(* IEC 61131-3 sources: volt/packages/volt-lsp-iec/test-corpus/CodesysTestProject/Device/Plc Logic/Application/Library Manager/Util, 115 files *)

(* ---- _STATE.dut ---- *)
TYPE _STATE :
(
	UNKNOWN := 0,
	DORMANT,
	STARTING,
	EXECUTING,
	CLEANING,
	DONE,
	ERROR,
	ABORTED,
	RESETTING
);
END_TYPE

(* ---- DATETIME.dut ---- *)
TYPE DATETIME :
STRUCT
	UIYEAR : YEAR;
	UIMONTH : MONTH;
	UIDAY : DAY;
	UIHOUR : HOUR;
	UIMINUTE : MINUTE;
	UISECOND : SECOND;
	UIMILLISECONDS : MILLISECOND;
	EWEEKDAY : WEEKDAY;
END_STRUCT
END_TYPE

(* ---- DAY.dut ---- *)
TYPE DAY : UINT (1..31);
END_TYPE

(* ---- DAYS.dut ---- *)
TYPE DAYS : BYTE;
END_TYPE

(* ---- ERROR.dut ---- *)
TYPE ERROR :
(
	_WRONG_TRANSITION := -1,
	_WRONG_CONFIGURATION := -2,
	NO_ERROR := 0,
	_TIME_OUT := 1,
	WRONG_CONFIGURATION := 2,
	RTC_HIGHRES_NOT_SUPPORTED,
	SYS_TIMEZONE_NOT_SUPPORTED
);
END_TYPE

(* ---- GEN_MODE.dut ---- *)
TYPE GEN_MODE :
(
	TRIANGLE := 0,
	TRIANGLE_POS := 1,
	SAWTOOTH_RISE := 2,
	SAWTOOTH_FALL := 3,
	RECTANGLE := 4,
	SINUS := 5,
	COSINUS := 6,
	SINE := 7,
	COSINE := 8
);
END_TYPE

(* ---- HOUR.dut ---- *)
TYPE HOUR : UINT (0..23);
END_TYPE

(* ---- MILLISECOND.dut ---- *)
TYPE MILLISECOND : UINT (0..999);
END_TYPE

(* ---- MINUTE.dut ---- *)
TYPE MINUTE : UINT (0..59);
END_TYPE

(* ---- MONTH.dut ---- *)
TYPE MONTH : UINT (1..12);
END_TYPE

(* ---- PERIOD.dut ---- *)
TYPE PERIOD :
(
	UNKNOWN := 0,
	STANDARD := 1,
	DAYLIGHT := 2
);
END_TYPE

(* ---- POINT.dut ---- *)
TYPE POINT :
STRUCT
	X : DINT;
	Y : DINT;
END_STRUCT
END_TYPE

(* ---- PT_SIZE.dut ---- *)
TYPE PT_SIZE :
STRUCT
	PSTRING : POINTER TO BYTE;
	UISIZE : UINT;
END_STRUCT
END_TYPE

(* ---- SCHEDULE.dut ---- *)
TYPE SCHEDULE :
STRUCT
	USISWITCH : USINT;
	TODFIRSTON : TIME_OF_DAY;
	TODLASTON : TIME_OF_DAY;
	BYDAYFLAGS : DAYS;
END_STRUCT
END_TYPE

(* ---- SECOND.dut ---- *)
TYPE SECOND : MINUTE;
END_TYPE

(* ---- SEGMENT.dut ---- *)
TYPE SEGMENT :
STRUCT
	SNAME : TZ_NAME;
	DTDATE : DateTime;
	IBIAS : INT;
END_STRUCT
END_TYPE

(* ---- TIMEZONE.dut ---- *)
TYPE TIMEZONE :
STRUCT
	IBIAS : INT;
	ASGPERIOD : ARRAY [1..2] OF Segment;
END_STRUCT
END_TYPE

(* ---- TZ_NAME.dut ---- *)
TYPE TZ_NAME : STRING(32);
END_TYPE

(* ---- WEEK.dut ---- *)
TYPE WEEK : UINT (1..53);
END_TYPE

(* ---- WEEKDAY.dut ---- *)
TYPE WEEKDAY :
(
	UNKNOWN := 0,
	MONDAY := 1,
	TUESDAY := 2,
	WEDNESDAY := 3,
	THURSDAY := 4,
	FRIDAY := 5,
	SATURDAY := 6,
	SUNDAY := 7
);
END_TYPE

(* ---- YEAR.dut ---- *)
TYPE YEAR : UINT (0..2106);
END_TYPE

(* ---- CONSTANTS.gvl ---- *)
VAR_GLOBAL
	GC_ULISECONDSINDAY : ULINT := (ANY_TO_ULINT(TIME#1440m0s0ms) / 1000);
	GC_AUSIWEEKDAY : ARRAY [0..11] OF USINT := [0, 3, 3, 6, 1, 4, 6, 2, 5, 0, 3, 5];
	GC_AUSIDAYSINMONTH : ARRAY [0..11] OF USINT := [31, 28, 31, 30, 31, 30, 31, 31, 30, 31, 30, 31];
	GC_AUIDAYSINYEAR : ARRAY [0..11] OF UINT := [0, 31, 59, 90, 120, 151, 181, 212, 243, 273, 304, 334];
	GC_DWSWITCHMASK : ARRAY [0..31] OF DWORD := [16#1, 16#2, 16#4, 16#8, 16#10, 16#20, 16#40, 16#80, 16#100, 16#200, 16#400, 16#800, 16#1000, 16#2000, 16#4000, 16#8000, 16#10000, 16#20000, 16#40000, 16#80000, 16#100000, 16#200000, 16#400000, 16#800000, 16#1000000, 16#2000000, 16#4000000, 16#8000000, 16#10000000, 16#20000000, 16#40000000, 16#80000000];
	GC_BYDAYMASK : ARRAY [0..7] OF DAYS := [DAY_FLAGS.EVERY_DAY, DAY_FLAGS.MONDAY, DAY_FLAGS.TUESDAY, DAY_FLAGS.WEDNESDAY, DAY_FLAGS.THURSDAY, DAY_FLAGS.FRIDAY, DAY_FLAGS.SATURDAY, DAY_FLAGS.SUNDAY];
END_VAR

(* ---- DAY_FLAGS.gvl ---- *)
VAR_GLOBAL
	EVERY_DAY : DAYS := 0;
	WORKING_DAYS : DAYS := 31;
	WEEKEND : DAYS := 96;
	MONDAY : DAYS := 1;
	TUESDAY : DAYS := 2;
	WEDNESDAY : DAYS := 4;
	THURSDAY : DAYS := 8;
	FRIDAY : DAYS := 16;
	SATURDAY : DAYS := 32;
	SUNDAY : DAYS := 64;
END_VAR

(* ---- GLOBALS.gvl ---- *)
VAR_GLOBAL
	G_DTPDATETIMEPROVIDER : DateTimeProvider;
END_VAR

(* ---- GVL_CONST.gvl ---- *)
VAR_GLOBAL
	UIBLOCKSIZEENCODED : UINT := REAL_TO_UINT((TextBlockSize.iBlockSize + (TextBlockSize.iBlockSize * 0.35)));
END_VAR

(* ---- TEXTBLOCKSIZE.gvl ---- *)
VAR_GLOBAL
	IBLOCKSIZE : INT := 22800;
END_VAR

(* ---- TSW.gvl ---- *)
VAR_GLOBAL
	GC_TZTIMEZONECET : TimeZone := STRUCT(iBias := 60, asgPeriod := [STRUCT(sName := 'CET', dtDate := STRUCT(uiMonth := 10, eWeekday := WEEKDAY.SUNDAY, uiDay := 5, uiHour := 3)), STRUCT(sName := 'CEST', dtDate := STRUCT(uiMonth := 3, eWeekday := WEEKDAY.SUNDAY, uiDay := 5, uiHour := 2), iBias := 60)]);
	GC_TZTIMEZONEUTC : TimeZone := STRUCT(asgPeriod := [STRUCT(sName := 'UTC')]);
END_VAR

(* ---- _IACTIONCONTROLLER.itf ---- *)
INTERFACE _IACTIONCONTROLLER
END_INTERFACE

METHOD CONTROLCLEANUPACTION
VAR_INPUT
	ITFCLEANUPACTIONPROVIDER : _ICleanupActionProvider;
	XABORTPROPOSED : BOOL;
	IERRORIDPROPOSED : INT;
END_VAR
VAR_OUTPUT
	XCOMPLETE : BOOL;
	XABORT : BOOL;
	IERRORID : INT;
END_VAR
END_METHOD

METHOD CONTROLCYCLICACTION
VAR_INPUT
	ITFCYCLICACTIONPROVIDER : _ICyclicActionProvider;
	ITFTIMINGCONTROLLER : _ITimingController;
END_VAR
VAR_OUTPUT
	XCOMPLETE : BOOL;
	IERRORID : INT;
END_VAR
END_METHOD

METHOD CONTROLEXITACTION
VAR_INPUT
	ITFEXITACTIONPROVIDER : _IExitActionProvider;
	XAFTERCLEANUP : BOOL;
	XINCOPYCODE : BOOL;
END_VAR
END_METHOD

METHOD CONTROLRESETACTION
VAR_INPUT
	ITFRESETACTIONPROVIDER : _IResetActionProvider;
END_VAR
VAR_OUTPUT
	XCOMPLETE : BOOL;
END_VAR
END_METHOD

METHOD CONTROLSTARTACTION
VAR_INPUT
	ITFSTARTACTIONPROVIDER : _IStartActionProvider;
END_VAR
VAR_OUTPUT
	XCOMPLETE : BOOL;
	IERRORID : INT;
END_VAR
END_METHOD

(* ---- _IACTIONPROVIDER.itf ---- *)
INTERFACE _IACTIONPROVIDER
END_INTERFACE

(* ---- _IBEHAVIOURMODEL.itf ---- *)
INTERFACE _IBEHAVIOURMODEL
END_INTERFACE

METHOD ABORTMODEL : ERROR
VAR_INPUT
	XCOMMIT : BOOL;
END_VAR
END_METHOD

METHOD GETMODELSTATE
VAR_INPUT
	XCOMMIT : BOOL;
END_VAR
VAR_OUTPUT
	XDONE : BOOL;
	XBUSY : BOOL;
	XERROR : BOOL;
	XABORTED : BOOL;
	IERRORID : INT;
	ESTATE : _STATE;
END_VAR
END_METHOD

METHOD RESETMODEL : ERROR
VAR_INPUT
	XCOMMIT : BOOL;
END_VAR
END_METHOD

METHOD STARTMODEL : ERROR
VAR_INPUT
	XCOMMIT : BOOL;
END_VAR
END_METHOD

(* ---- _ICLEANUPACTIONPROVIDER.itf ---- *)
INTERFACE _ICLEANUPACTIONPROVIDER
END_INTERFACE

METHOD CLEANUPACTION
VAR_INPUT
	XABORTPROPOSED : BOOL;
	IERRORIDPROPOSED : INT;
END_VAR
VAR_OUTPUT
	XCOMPLETE : BOOL;
	XABORT : BOOL;
	IERRORID : INT;
END_VAR
END_METHOD

(* ---- _ICONFIGURATIONPROVIDER.itf ---- *)
INTERFACE _ICONFIGURATIONPROVIDER
END_INTERFACE

METHOD GETCONFIGURATION
VAR_OUTPUT
	XLEVELCONTROLLED : BOOL;
	XTIMINGCONTROLLED : BOOL;
	XTIMELIMITED : BOOL;
	XTIMEOUTCONSTRAINT : BOOL;
	XABORTABLE : BOOL;
	XEDGETRIGGERED : BOOL;
	XHASCONTINUOUSBEHAVIOUR : BOOL;
	XSUPPORTSEXITACTION : BOOL;
END_VAR
END_METHOD

(* ---- _ICONFIGURATIONPROVIDER2.itf ---- *)
INTERFACE _ICONFIGURATIONPROVIDER2
END_INTERFACE

METHOD GETCONFIGURATION2
VAR_OUTPUT
	XLEVELCONTROLLED : BOOL;
	XTIMINGCONTROLLED : BOOL;
	XTIMELIMITED : BOOL;
	XTIMEOUTCONSTRAINT : BOOL;
	XABORTABLE : BOOL;
	XEDGETRIGGERED : BOOL;
	XHASCONTINUOUSBEHAVIOUR : BOOL;
	XSUPPORTSEXITACTION : BOOL;
	XSUPPORTSSAMPLEACTION : BOOL;
END_VAR
END_METHOD

(* ---- _ICYCLICACTIONPROVIDER.itf ---- *)
INTERFACE _ICYCLICACTIONPROVIDER
END_INTERFACE

METHOD CYCLICACTION
VAR_INPUT
	ITFTIMINGCONTROLLER : _ITimingController;
END_VAR
VAR_OUTPUT
	XCOMPLETE : BOOL;
	IERRORID : INT;
END_VAR
END_METHOD

(* ---- _IEXITACTIONPROVIDER.itf ---- *)
INTERFACE _IEXITACTIONPROVIDER
END_INTERFACE

METHOD EXITACTION
VAR_INPUT
	XAFTERCLEANUP : BOOL;
	XINCOPYCODE : BOOL;
END_VAR
END_METHOD

(* ---- _IHASCONTINUOUSBEHAVIOUR.itf ---- *)
INTERFACE _IHASCONTINUOUSBEHAVIOUR
END_INTERFACE

(* ---- _ILEVELCONTROLLED.itf ---- *)
INTERFACE _ILEVELCONTROLLED
END_INTERFACE

(* ---- _IRESETACTIONPROVIDER.itf ---- *)
INTERFACE _IRESETACTIONPROVIDER
END_INTERFACE

METHOD RESETACTION
VAR_OUTPUT
	XCOMPLETE : BOOL;
END_VAR
END_METHOD

(* ---- _ISTARTACTIONPROVIDER.itf ---- *)
INTERFACE _ISTARTACTIONPROVIDER
END_INTERFACE

METHOD STARTACTION
VAR_OUTPUT
	XCOMPLETE : BOOL;
	IERRORID : INT;
END_VAR
END_METHOD

(* ---- _ITIMINGCONTROLLER.itf ---- *)
INTERFACE _ITIMINGCONTROLLER
END_INTERFACE

METHOD CONTROLLERCHECKTIMING
VAR_OUTPUT
	XTIMEOUT : BOOL;
	XTIMELIMIT : BOOL;
END_VAR
END_METHOD

METHOD STARTINVOCATIONTIMER
END_METHOD

METHOD STARTOPERATIONTIMER
END_METHOD

(* ---- IDATETIMEPROVIDER.itf ---- *)
INTERFACE IDATETIMEPROVIDER
END_INTERFACE

METHOD GETDATETIME : ULINT
VAR_OUTPUT
	EERRORID : ERROR;
END_VAR
END_METHOD

(* ---- ITIMESWITCH.itf ---- *)
INTERFACE ITIMESWITCH
END_INTERFACE

(* ---- BASE64.pou ---- *)
FUNCTION BASE64 : PT_SIZE
VAR_INPUT
	TEXTTOENCODE : PT_SIZE;
	ISLASTBLOCK : BOOL;
	PBYERROR : POINTER TO BYTE;
END_VAR
END_FUNCTION

(* ---- BCD_TO_BYTE.pou ---- *)
FUNCTION BCD_TO_BYTE : BYTE
VAR_INPUT
	B : BYTE;
END_VAR
END_FUNCTION

(* ---- BCD_TO_DWORD.pou ---- *)
FUNCTION BCD_TO_DWORD : DWORD
VAR_INPUT
	X : DWORD;
END_VAR
END_FUNCTION

(* ---- BCD_TO_INT.pou ---- *)
FUNCTION BCD_TO_INT : INT
VAR_INPUT
	B : BYTE;
END_VAR
END_FUNCTION

(* ---- BCD_TO_WORD.pou ---- *)
FUNCTION BCD_TO_WORD : WORD
VAR_INPUT
	W : WORD;
END_VAR
END_FUNCTION

(* ---- BYTE_TO_BCD.pou ---- *)
FUNCTION BYTE_TO_BCD : BYTE
VAR_INPUT
	B : BYTE;
END_VAR
END_FUNCTION

(* ---- BYTE_TO_GRAY.pou ---- *)
FUNCTION BYTE_TO_GRAY : BYTE
VAR_INPUT
	B : BYTE;
END_VAR
END_FUNCTION

(* ---- BYTE_TO_HEXINASCII.pou ---- *)
FUNCTION BYTE_TO_HEXINASCII : WORD
VAR_INPUT
	B : BYTE;
END_VAR
END_FUNCTION

(* ---- COMBINEDATETIME.pou ---- *)
FUNCTION COMBINEDATETIME : ULINT
VAR_INPUT
	DATDATE : DATE;
	TODTIME : TIME_OF_DAY;
END_VAR
VAR_OUTPUT
	EERRORID : ERROR := ERROR.NO_ERROR;
END_VAR
END_FUNCTION

(* ---- CONVERTDATETIME.pou ---- *)
FUNCTION CONVERTDATETIME : ULINT
VAR_INPUT
	UIYEAR : YEAR;
END_VAR
VAR_OUTPUT
	EERRORID : ERROR;
END_VAR
VAR_IN_OUT
	DTDATETIME : DateTime;
END_VAR
END_FUNCTION

(* ---- DATETIMEFROMWEEK.pou ---- *)
FUNCTION DATETIMEFROMWEEK : ULINT
VAR_INPUT
	UIYEAR : YEAR;
	UIWEEK : WEEK;
	EWEEKDAY : WEEKDAY;
END_VAR
VAR_OUTPUT
	EERRORID : ERROR;
END_VAR
END_FUNCTION

(* ---- DAYOFWEEK.pou ---- *)
FUNCTION DAYOFWEEK : WEEKDAY
VAR_INPUT
	DATDATE : DATE;
END_VAR
VAR_OUTPUT
	EERRORID : ERROR := ERROR.NO_ERROR;
END_VAR
END_FUNCTION

(* ---- DWORD_TO_BCD.pou ---- *)
FUNCTION DWORD_TO_BCD : DWORD
VAR_INPUT
	X : DWORD;
END_VAR
END_FUNCTION

(* ---- DWORD_TO_GRAY.pou ---- *)
FUNCTION DWORD_TO_GRAY : DWORD
VAR_INPUT
	X : DWORD;
END_VAR
END_FUNCTION

(* ---- EXTRACT.pou ---- *)
FUNCTION EXTRACT : BOOL
VAR_INPUT
	X : DWORD;
	N : BYTE;
END_VAR
END_FUNCTION

(* ---- EXTRACTYEARMONTHDAY.pou ---- *)
FUNCTION EXTRACTYEARMONTHDAY : ERROR
VAR_INPUT
	ULIDATETIME : ULINT;
END_VAR
VAR_OUTPUT
	UIYEAR : YEAR;
	UIMONTH : MONTH;
	UIDAY : DAY;
END_VAR
END_FUNCTION

(* ---- GETBIT.pou ---- *)
FUNCTION GETBIT : BOOL
VAR_INPUT
	X : LWORD;
	N : BYTE;
END_VAR
END_FUNCTION

(* ---- GETDATETIME.pou ---- *)
FUNCTION GETDATETIME : ULINT
VAR_OUTPUT
	EERRORID : ERROR;
END_VAR
END_FUNCTION

(* ---- GETLIBVERSION.pou ---- *)
FUNCTION GETLIBVERSION : VERSION
END_FUNCTION

(* ---- GETLIBVERSIONNUMBER.pou ---- *)
FUNCTION GETLIBVERSIONNUMBER : DWORD
END_FUNCTION

(* ---- GETLOCALDATETIME.pou ---- *)
FUNCTION GETLOCALDATETIME : ULINT
VAR_OUTPUT
	EERRORID : ERROR;
END_VAR
VAR_IN_OUT
	TZTIMEZONE : TimeZone;
END_VAR
END_FUNCTION

(* ---- GETTIMESTAMPSDIFFERENCE.pou ---- *)
FUNCTION GETTIMESTAMPSDIFFERENCE : ERROR
VAR_INPUT
	ULIDATETIMEFIRST : ULINT;
	ULIDATETIMESECOND : ULINT;
END_VAR
VAR_OUTPUT
	ULIDAYS : ULINT;
	UIHOURS : HOUR;
	UIMINUTES : MINUTE;
	UISECONDS : SECOND;
	UIMILLISECONDS : MILLISECOND;
END_VAR
END_FUNCTION

(* ---- GRAY_TO_BYTE.pou ---- *)
FUNCTION GRAY_TO_BYTE : BYTE
VAR_INPUT
	B : BYTE;
END_VAR
END_FUNCTION

(* ---- GRAY_TO_DWORD.pou ---- *)
FUNCTION GRAY_TO_DWORD : DWORD
VAR_INPUT
	X : DWORD;
END_VAR
END_FUNCTION

(* ---- GRAY_TO_WORD.pou ---- *)
FUNCTION GRAY_TO_WORD : WORD
VAR_INPUT
	W : WORD;
END_VAR
END_FUNCTION

(* ---- HEXINASCII_TO_BYTE.pou ---- *)
FUNCTION HEXINASCII_TO_BYTE : BYTE
VAR_INPUT
	W : WORD;
END_VAR
END_FUNCTION

(* ---- INT_TO_BCD.pou ---- *)
FUNCTION INT_TO_BCD : BYTE
VAR_INPUT
	I : INT;
END_VAR
END_FUNCTION

(* ---- ISLEAPYEAR.pou ---- *)
FUNCTION ISLEAPYEAR : BOOL
VAR_INPUT
	UIYEAR : YEAR;
END_VAR
VAR_OUTPUT
	EERRORID : ERROR := ERROR.NO_ERROR;
END_VAR
END_FUNCTION

(* ---- ISLIBRELEASED.pou ---- *)
FUNCTION ISLIBRELEASED : BOOL
END_FUNCTION

(* ---- JOINDATETIME.pou ---- *)
FUNCTION JOINDATETIME : ULINT
VAR_INPUT
	UIYEAR : YEAR;
	UIMONTH : MONTH;
	UIDAY : DAY;
	UIHOUR : HOUR;
	UIMINUTE : MINUTE;
	UISECOND : SECOND;
	UIMILLISECONDS : MILLISECOND;
END_VAR
VAR_OUTPUT
	EERRORID : ERROR := ERROR.NO_ERROR;
END_VAR
END_FUNCTION

(* ---- JOINYEARMONTHDAY.pou ---- *)
FUNCTION JOINYEARMONTHDAY : ULINT
VAR_INPUT
	UIYEAR : YEAR;
	UIMONTH : MONTH;
	UIDAY : DAY;
END_VAR
VAR_OUTPUT
	EERRORID : ERROR := ERROR.NO_ERROR;
END_VAR
END_FUNCTION

(* ---- LASTWEEKOFYEAR.pou ---- *)
FUNCTION LASTWEEKOFYEAR : Week
VAR_INPUT
	UIYEAR : YEAR;
END_VAR
VAR_OUTPUT
	EERRORID : ERROR;
END_VAR
END_FUNCTION

(* ---- LEAPYEARS.pou ---- *)
FUNCTION LEAPYEARS : UINT
VAR_INPUT
	UISTARTYEAR : YEAR;
	UIENDYEAR : YEAR;
END_VAR
VAR_OUTPUT
	EERRORID : ERROR;
END_VAR
END_FUNCTION

(* ---- LOCALDATETIME.pou ---- *)
FUNCTION LOCALDATETIME : ULINT
VAR_INPUT
	ULIDATETIME : ULINT;
END_VAR
VAR_OUTPUT
	EERRORID : ERROR;
	EPERIOD : PERIOD;
END_VAR
VAR_IN_OUT
	TZTIMEZONE : TimeZone;
END_VAR
END_FUNCTION

(* ---- PACK.pou ---- *)
FUNCTION PACK : BYTE
VAR_INPUT
	B0 : BOOL;
	B1 : BOOL;
	B2 : BOOL;
	B3 : BOOL;
	B4 : BOOL;
	B5 : BOOL;
	B6 : BOOL;
	B7 : BOOL;
END_VAR
END_FUNCTION

(* ---- PUTBIT.pou ---- *)
FUNCTION PUTBIT : DWORD
VAR_INPUT
	X : DWORD;
	N : BYTE;
	B : BOOL;
END_VAR
END_FUNCTION

(* ---- SEPARATEDATETIME.pou ---- *)
FUNCTION SEPARATEDATETIME : ERROR
VAR_INPUT
	ULIDATETIME : ULINT;
END_VAR
VAR_OUTPUT
	EWEEKDAY : WEEKDAY;
	DATDATE : DATE;
	TODTIME : TIME_OF_DAY;
END_VAR
END_FUNCTION

(* ---- SETBIT.pou ---- *)
FUNCTION SETBIT : BOOL
VAR_INPUT
	X : __SYSTEM.AnyType;
	N : BYTE;
	B : BOOL;
END_VAR
END_FUNCTION

(* ---- SPLITDATETIME.pou ---- *)
FUNCTION SPLITDATETIME : ERROR
VAR_INPUT
	ULIDATETIME : ULINT;
END_VAR
VAR_OUTPUT
	UIYEAR : YEAR;
	UIMONTH : MONTH;
	UIDAY : DAY;
	UIHOUR : HOUR;
	UIMINUTE : MINUTE;
	UISECOND : SECOND;
	UIMILLISECONDS : MILLISECOND;
	EWEEKDAY : WEEKDAY;
END_VAR
END_FUNCTION

(* ---- SWITCHBIT.pou ---- *)
FUNCTION SWITCHBIT : DWORD
VAR_INPUT
	X : DWORD;
	N : BYTE;
END_VAR
END_FUNCTION

(* ---- WEEKOFYEAR.pou ---- *)
FUNCTION WEEKOFYEAR : ERROR
VAR_INPUT
	ULIDATETIME : ULINT;
END_VAR
VAR_OUTPUT
	UIYEAR : YEAR;
	UIWEEK : WEEK;
	EWEEKDAY : WEEKDAY;
END_VAR
END_FUNCTION

(* ---- WORD_AS_STRING.pou ---- *)
FUNCTION WORD_AS_STRING : STRING(2)
VAR_INPUT
	W : WORD;
	ORDER : BOOL;
END_VAR
END_FUNCTION

(* ---- WORD_TO_BCD.pou ---- *)
FUNCTION WORD_TO_BCD : WORD
VAR_INPUT
	W : WORD;
END_VAR
END_FUNCTION

(* ---- WORD_TO_GRAY.pou ---- *)
FUNCTION WORD_TO_GRAY : WORD
VAR_INPUT
	W : WORD;
END_VAR
END_FUNCTION

(* ---- _BEHAVIOURMODEL.pou ---- *)
FUNCTION_BLOCK _BEHAVIOURMODEL
VAR_INPUT
	ITFACTIONPROVIDER : _IActionProvider;
	ITFTIMINGCONTROLLER : _ITimingController;
	XCONTROL : BOOL;
	XABORT : BOOL;
	UDITIMELIMIT : UDINT;
	UDITIMEOUT : UDINT;
END_VAR
VAR_OUTPUT
	XDONE : BOOL;
	XBUSY : BOOL;
	XERROR : BOOL;
	XABORTED : BOOL;
	IERRORID : INT;
	ESTATE : _STATE;
	EINTERNALERRORID : ERROR;
END_VAR
VAR
	_ITFACTIONPROVIDER : _IActionProvider;
	_ITFACTIONCONTROLLER : _IActionController;
	_XLEVELCONTROLLED : BOOL;
	_XTIMINGCONTROLLED : BOOL;
	_XTIMELIMITED : BOOL;
	_XTIMEOUTCONSTRAINT : BOOL;
	_XABORTABLE : BOOL;
	_XEDGETRIGGERED : BOOL;
	_XHASCONTINUOUSBEHAVIOUR : BOOL;
	_XSUPPORTSEXITACTION : BOOL;
	_XSUPPORTSSAMPLEACTION : BOOL;
	_XRESETREQUEST : BOOL;
	_XABORTPROPOSED : BOOL;
	_IERRORIDPROPOSED : INT;
	_XFIRSTHANDLESTARTINGSTATECALL : BOOL;
	_XLASTAGAIN : BOOL;
	_ITFSTARTACTIONPROVIDER : _IStartActionProvider;
	_ITFCYCLICACTIONPROVIDER : _ICyclicActionProvider;
	_ITFCLEANUPACTIONPROVIDER : _ICleanupActionProvider;
	_ITFEXITACTIONPROVIDER : _IExitActionProvider;
	_ITFRESETACTIONPROVIDER : _IResetActionProvider;
	ACTIONCONTROLLER : _IActionController;
	MODELTIMELIMIT : UDINT;
	MODELTIMEOUT : UDINT;
END_VAR
END_FUNCTION_BLOCK

METHOD _CHECKABORTCONDITION : BOOL
END_METHOD

METHOD _CHECKPARAMETER
VAR_OUTPUT
	EERRORID : ERROR;
END_VAR
END_METHOD

METHOD _CHECKTIMEOUTCONDITION
END_METHOD

METHOD _EXECUTE
VAR_OUTPUT
	EERRORID : ERROR := ERROR.NO_ERROR;
END_VAR
END_METHOD

METHOD _RESETACTION
END_METHOD

METHOD ABORTMODEL : ERROR
VAR_INPUT
	XCOMMIT : BOOL;
END_VAR
END_METHOD

METHOD GETCONFIGURATION
VAR_OUTPUT
	XLEVELCONTROLLED : BOOL;
	XTIMINGCONTROLLED : BOOL;
	XTIMELIMITED : BOOL;
	XTIMEOUTCONSTRAINT : BOOL;
	XABORTABLE : BOOL;
	XEDGETRIGGERED : BOOL;
	XHASCONTINUOUSBEHAVIOUR : BOOL;
	XSUPPORTSEXITACTION : BOOL;
END_VAR
END_METHOD

METHOD GETCONFIGURATION2
VAR_OUTPUT
	XLEVELCONTROLLED : BOOL;
	XTIMINGCONTROLLED : BOOL;
	XTIMELIMITED : BOOL;
	XTIMEOUTCONSTRAINT : BOOL;
	XABORTABLE : BOOL;
	XEDGETRIGGERED : BOOL;
	XHASCONTINUOUSBEHAVIOUR : BOOL;
	XSUPPORTSEXITACTION : BOOL;
	XSUPPORTSSAMPLEACTION : BOOL;
END_VAR
END_METHOD

METHOD GETMODELSTATE
VAR_INPUT
	XCOMMIT : BOOL;
END_VAR
VAR_OUTPUT
	XDONE : BOOL;
	XBUSY : BOOL;
	XERROR : BOOL;
	XABORTED : BOOL;
	IERRORID : INT;
	ESTATE : _STATE;
END_VAR
END_METHOD

METHOD RESETMODEL : ERROR
VAR_INPUT
	XCOMMIT : BOOL;
END_VAR
END_METHOD

METHOD STARTMODEL : ERROR
VAR_INPUT
	XCOMMIT : BOOL;
END_VAR
END_METHOD

METHOD _HANDLEABORTEDSTATE
VAR_OUTPUT
	XAGAIN : BOOL;
END_VAR
END_METHOD

METHOD _HANDLECLEANINGSTATE
VAR_OUTPUT
	XAGAIN : BOOL;
END_VAR
END_METHOD

METHOD _HANDLEDONESTATE
VAR_OUTPUT
	XAGAIN : BOOL;
END_VAR
END_METHOD

METHOD _HANDLEDORMANTSTATE
VAR_OUTPUT
	XAGAIN : BOOL;
END_VAR
END_METHOD

METHOD _HANDLEERRORSTATE
VAR_OUTPUT
	XAGAIN : BOOL;
END_VAR
END_METHOD

METHOD _HANDLEEXECUTINGSTATE
VAR_OUTPUT
	XAGAIN : BOOL;
END_VAR
END_METHOD

METHOD _HANDLERESETTINGSTATE
VAR_OUTPUT
	XAGAIN : BOOL;
END_VAR
END_METHOD

METHOD _HANDLESTARTINGSTATE
VAR_OUTPUT
	XAGAIN : BOOL;
	IERRORID : INT;
END_VAR
END_METHOD

METHOD _STATEMACHINE : ERROR
END_METHOD

(* ---- _LCONC.pou ---- *)
FUNCTION_BLOCK _LCONC
VAR_INPUT
	XENABLE : BOOL;
END_VAR
VAR_OUTPUT
	XBUSY : BOOL;
	XERROR : BOOL;
END_VAR
VAR
	_MODEL : _BehaviourModel := STRUCT(itfActionProvider := THIS^, itfTimingController := 0);
	ACTIONCONTROLLER : _IActionController;
	MODELTIMELIMIT : UDINT;
	MODELTIMEOUT : UDINT;
END_VAR
END_FUNCTION_BLOCK

METHOD FB_EXIT : BOOL
VAR_INPUT
	BINCOPYCODE : BOOL;
END_VAR
END_METHOD

METHOD _EXECUTE
VAR_OUTPUT
	EERRORID : ERROR;
END_VAR
END_METHOD

METHOD CLEANUPACTION
VAR_INPUT
	XABORTPROPOSED : BOOL;
	IERRORIDPROPOSED : INT;
END_VAR
VAR_OUTPUT
	XCOMPLETE : BOOL := TRUE;
	XABORT : BOOL := xAbortProposed;
	IERRORID : INT := iErrorIDProposed;
END_VAR
END_METHOD

METHOD CYCLICACTION
VAR_INPUT
	ITFTIMINGCONTROLLER : _ITimingController;
END_VAR
VAR_OUTPUT
	XCOMPLETE : BOOL := TRUE;
	IERRORID : INT := 0;
END_VAR
END_METHOD

METHOD EXITACTION
VAR_INPUT
	XAFTERCLEANUP : BOOL;
	XINCOPYCODE : BOOL;
END_VAR
END_METHOD

METHOD RESETACTION
VAR_OUTPUT
	XCOMPLETE : BOOL := TRUE;
END_VAR
END_METHOD

METHOD STARTACTION
VAR_OUTPUT
	XCOMPLETE : BOOL := TRUE;
	IERRORID : INT := 0;
END_VAR
END_METHOD

METHOD ABORTMODEL : ERROR
VAR_INPUT
	XCOMMIT : BOOL;
END_VAR
END_METHOD

METHOD GETCONFIGURATION
VAR_OUTPUT
	XLEVELCONTROLLED : BOOL;
	XTIMINGCONTROLLED : BOOL;
	XTIMELIMITED : BOOL;
	XTIMEOUTCONSTRAINT : BOOL;
	XABORTABLE : BOOL;
	XEDGETRIGGERED : BOOL;
	XHASCONTINUOUSBEHAVIOUR : BOOL;
	XSUPPORTSEXITACTION : BOOL;
END_VAR
END_METHOD

METHOD GETCONFIGURATION2
VAR_OUTPUT
	XLEVELCONTROLLED : BOOL;
	XTIMINGCONTROLLED : BOOL;
	XTIMELIMITED : BOOL;
	XTIMEOUTCONSTRAINT : BOOL;
	XABORTABLE : BOOL;
	XEDGETRIGGERED : BOOL;
	XHASCONTINUOUSBEHAVIOUR : BOOL;
	XSUPPORTSEXITACTION : BOOL;
	XSUPPORTSSAMPLEACTION : BOOL;
END_VAR
END_METHOD

METHOD GETMODELSTATE
VAR_INPUT
	XCOMMIT : BOOL;
END_VAR
VAR_OUTPUT
	XDONE : BOOL;
	XBUSY : BOOL;
	XERROR : BOOL;
	XABORTED : BOOL;
	IERRORID : INT;
	ESTATE : _STATE;
END_VAR
END_METHOD

METHOD RESETMODEL : ERROR
VAR_INPUT
	XCOMMIT : BOOL;
END_VAR
END_METHOD

METHOD STARTMODEL : ERROR
VAR_INPUT
	XCOMMIT : BOOL;
END_VAR
END_METHOD

(* ---- BIT_AS_BYTE.pou ---- *)
FUNCTION_BLOCK BIT_AS_BYTE
VAR_INPUT
	B0 : BOOL;
	B1 : BOOL;
	B2 : BOOL;
	B3 : BOOL;
	B4 : BOOL;
	B5 : BOOL;
	B6 : BOOL;
	B7 : BOOL;
END_VAR
VAR_OUTPUT
	B : BYTE;
END_VAR
END_FUNCTION_BLOCK

(* ---- BIT_AS_DWORD.pou ---- *)
FUNCTION_BLOCK BIT_AS_DWORD
VAR_INPUT
	B00 : BOOL;
	B01 : BOOL;
	B02 : BOOL;
	B03 : BOOL;
	B04 : BOOL;
	B05 : BOOL;
	B06 : BOOL;
	B07 : BOOL;
	B08 : BOOL;
	B09 : BOOL;
	B10 : BOOL;
	B11 : BOOL;
	B12 : BOOL;
	B13 : BOOL;
	B14 : BOOL;
	B15 : BOOL;
	B16 : BOOL;
	B17 : BOOL;
	B18 : BOOL;
	B19 : BOOL;
	B20 : BOOL;
	B21 : BOOL;
	B22 : BOOL;
	B23 : BOOL;
	B24 : BOOL;
	B25 : BOOL;
	B26 : BOOL;
	B27 : BOOL;
	B28 : BOOL;
	B29 : BOOL;
	B30 : BOOL;
	B31 : BOOL;
END_VAR
VAR_OUTPUT
	X : DWORD;
END_VAR
END_FUNCTION_BLOCK

(* ---- BIT_AS_WORD.pou ---- *)
FUNCTION_BLOCK BIT_AS_WORD
VAR_INPUT
	B00 : BOOL;
	B01 : BOOL;
	B02 : BOOL;
	B03 : BOOL;
	B04 : BOOL;
	B05 : BOOL;
	B06 : BOOL;
	B07 : BOOL;
	B08 : BOOL;
	B09 : BOOL;
	B10 : BOOL;
	B11 : BOOL;
	B12 : BOOL;
	B13 : BOOL;
	B14 : BOOL;
	B15 : BOOL;
END_VAR
VAR_OUTPUT
	W : WORD;
END_VAR
END_FUNCTION_BLOCK

(* ---- BLINK.pou ---- *)
FUNCTION_BLOCK BLINK
VAR_INPUT
	ENABLE : BOOL;
	TIMELOW : TIME;
	TIMEHIGH : TIME;
END_VAR
VAR_OUTPUT
	OUT : BOOL;
END_VAR
VAR
	CLOCK : TP;
END_VAR
END_FUNCTION_BLOCK

(* ---- BYTE_AS_BIT.pou ---- *)
FUNCTION_BLOCK BYTE_AS_BIT
VAR_INPUT
	B : BYTE;
END_VAR
VAR_OUTPUT
	B0 : BOOL;
	B1 : BOOL;
	B2 : BOOL;
	B3 : BOOL;
	B4 : BOOL;
	B5 : BOOL;
	B6 : BOOL;
	B7 : BOOL;
END_VAR
END_FUNCTION_BLOCK

(* ---- CHARCURVE.pou ---- *)
FUNCTION_BLOCK CHARCURVE
VAR_INPUT
	IN : INT;
	N : BYTE;
END_VAR
VAR_OUTPUT
	OUT : INT;
	ERR : BYTE;
END_VAR
VAR_IN_OUT
	P : ARRAY [0..10] OF POINT;
END_VAR
VAR
	I : INT;
END_VAR
END_FUNCTION_BLOCK

(* ---- DATETIMEPROVIDER.pou ---- *)
FUNCTION_BLOCK DATETIMEPROVIDER
END_FUNCTION_BLOCK

METHOD GETDATETIME : ULINT
VAR_OUTPUT
	EERRORID : ERROR;
END_VAR
END_METHOD

(* ---- DERIVATIVE.pou ---- *)
FUNCTION_BLOCK DERIVATIVE
VAR_INPUT
	IN : REAL;
	TM : DWORD;
	RESET : BOOL;
END_VAR
VAR_OUTPUT
	OUT : REAL;
END_VAR
VAR
	X3 : REAL;
	X2 : REAL;
	X1 : REAL;
	T2 : DWORD;
	T1 : DWORD;
	_INIT : BOOL := TRUE;
END_VAR
END_FUNCTION_BLOCK

(* ---- DWORD_AS_BIT.pou ---- *)
FUNCTION_BLOCK DWORD_AS_BIT
VAR_INPUT
	X : DWORD;
END_VAR
VAR_OUTPUT
	B00 : BOOL;
	B01 : BOOL;
	B02 : BOOL;
	B03 : BOOL;
	B04 : BOOL;
	B05 : BOOL;
	B06 : BOOL;
	B07 : BOOL;
	B08 : BOOL;
	B09 : BOOL;
	B10 : BOOL;
	B11 : BOOL;
	B12 : BOOL;
	B13 : BOOL;
	B14 : BOOL;
	B15 : BOOL;
	B16 : BOOL;
	B17 : BOOL;
	B18 : BOOL;
	B19 : BOOL;
	B20 : BOOL;
	B21 : BOOL;
	B22 : BOOL;
	B23 : BOOL;
	B24 : BOOL;
	B25 : BOOL;
	B26 : BOOL;
	B27 : BOOL;
	B28 : BOOL;
	B29 : BOOL;
	B30 : BOOL;
	B31 : BOOL;
END_VAR
END_FUNCTION_BLOCK

(* ---- FREQ_MEASURE.pou ---- *)
FUNCTION_BLOCK FREQ_MEASURE
VAR_INPUT
	IN : BOOL;
	PERIODS : INT (1..10) := 1;
	RESET : BOOL;
END_VAR
VAR_OUTPUT
	OUT : REAL;
	VALID : BOOL;
END_VAR
VAR
	OLDIN : BOOL;
	_INIT : BOOL;
	OLDT : TIME;
	DIFF : DWORD;
	ADIFF : ARRAY [0..9] OF DWORD;
	V : INT;
	B : INT;
	I : INT;
END_VAR
END_FUNCTION_BLOCK

(* ---- GEN.pou ---- *)
FUNCTION_BLOCK GEN
VAR_INPUT
	MODE : GEN_MODE;
	BASE : BOOL;
	PERIOD : TIME := TIME#1s0ms;
	CYCLES : INT := 1000;
	AMPLITUDE : INT;
	RESET : BOOL;
END_VAR
VAR_OUTPUT
	OUT : INT;
END_VAR
VAR
	CET : DINT;
	PER : DINT;
	COUNTER : INT;
	CLOCK : TON;
END_VAR
END_FUNCTION_BLOCK

(* ---- HYSTERESIS.pou ---- *)
FUNCTION_BLOCK HYSTERESIS
VAR_INPUT
	IN : INT;
	HIGH : INT;
	LOW : INT;
END_VAR
VAR_OUTPUT
	OUT : BOOL;
END_VAR
END_FUNCTION_BLOCK

(* ---- INTEGRAL.pou ---- *)
FUNCTION_BLOCK INTEGRAL
VAR_INPUT
	IN : REAL;
	TM : DWORD;
	RESET : BOOL;
END_VAR
VAR_OUTPUT
	OUT : REAL;
	OVERFLOW : BOOL := FALSE;
END_VAR
END_FUNCTION_BLOCK

(* ---- LIMITALARM.pou ---- *)
FUNCTION_BLOCK LIMITALARM
VAR_INPUT
	IN : INT;
	HIGH : INT;
	LOW : INT;
END_VAR
VAR_OUTPUT
	O : BOOL;
	U : BOOL;
	IL : BOOL;
END_VAR
END_FUNCTION_BLOCK

(* ---- LIN_TRAFO.pou ---- *)
FUNCTION_BLOCK LIN_TRAFO
VAR_INPUT
	IN : REAL;
	IN_MIN : REAL;
	IN_MAX : REAL;
	OUT_MIN : REAL;
	OUT_MAX : REAL;
END_VAR
VAR_OUTPUT
	OUT : REAL;
	ERROR : BOOL;
END_VAR
VAR
	DIFF : REAL;
END_VAR
END_FUNCTION_BLOCK

(* ---- PD.pou ---- *)
FUNCTION_BLOCK PD
VAR_INPUT
	ACTUAL : REAL;
	SET_POINT : REAL;
	KP : REAL;
	TV : REAL;
	Y_MANUAL : REAL;
	Y_OFFSET : REAL;
	Y_MIN : REAL;
	Y_MAX : REAL;
	MANUAL : BOOL;
	RESET : BOOL;
END_VAR
VAR_OUTPUT
	Y : REAL;
	LIMITS_ACTIVE : BOOL := FALSE;
END_VAR
VAR
	CLOCK : TON;
	D : DERIVATIVE;
	TMDIFF : DWORD;
	ERROR : REAL;
	_INIT : BOOL := TRUE;
	Y_ADDOFFSET : REAL;
	KPCOPY : REAL;
	TVCOPY : REAL;
END_VAR
END_FUNCTION_BLOCK

(* ---- PID.pou ---- *)
FUNCTION_BLOCK PID
VAR_INPUT
	ACTUAL : REAL;
	SET_POINT : REAL;
	KP : REAL;
	TN : REAL;
	TV : REAL;
	Y_MANUAL : REAL;
	Y_OFFSET : REAL;
	Y_MIN : REAL;
	Y_MAX : REAL;
	MANUAL : BOOL;
	RESET : BOOL;
END_VAR
VAR_OUTPUT
	Y : REAL;
	LIMITS_ACTIVE : BOOL := FALSE;
	OVERFLOW : BOOL := FALSE;
END_VAR
VAR
	CLOCK : TON;
	I : INTEGRAL;
	D : DERIVATIVE;
	TMDIFF : DWORD;
	ERROR : REAL;
	_INIT : BOOL := TRUE;
	Y_ADDOFFSET : REAL;
	KPCOPY : REAL;
	TNCOPY : REAL;
	TVCOPY : REAL;
END_VAR
END_FUNCTION_BLOCK

(* ---- PID_FIXCYCLE.pou ---- *)
FUNCTION_BLOCK PID_FIXCYCLE
VAR_INPUT
	ACTUAL : REAL;
	SET_POINT : REAL;
	KP : REAL;
	TN : REAL;
	TV : REAL;
	Y_MANUAL : REAL;
	Y_OFFSET : REAL;
	Y_MIN : REAL;
	Y_MAX : REAL;
	MANUAL : BOOL;
	RESET : BOOL;
	CYCLE : REAL;
END_VAR
VAR_OUTPUT
	Y : REAL;
	LIMITS_ACTIVE : BOOL := FALSE;
	OVERFLOW : BOOL := FALSE;
END_VAR
VAR
	I : INTEGRAL;
	D : DERIVATIVE;
	TMDIFF : DWORD;
	ERROR : REAL;
	_INIT : BOOL := TRUE;
	Y_ADDOFFSET : REAL;
	KPCOPY : REAL;
	TNCOPY : REAL;
	TVCOPY : REAL;
END_VAR
END_FUNCTION_BLOCK

(* ---- RAMP_INT.pou ---- *)
FUNCTION_BLOCK RAMP_INT
VAR_INPUT
	IN : INT;
	ASCEND : INT;
	DESCEND : INT;
	TIMEBASE : TIME;
	RESET : BOOL;
END_VAR
VAR_OUTPUT
	OUT : INT;
END_VAR
VAR
	DIFF : DINT;
	OLD_IN : INT;
	TB : DWORD;
	CET : DWORD;
	CH : INT;
	CLOCK : TON;
END_VAR
END_FUNCTION_BLOCK

(* ---- RAMP_REAL.pou ---- *)
FUNCTION_BLOCK RAMP_REAL
VAR_INPUT
	IN : REAL;
	ASCEND : REAL;
	DESCEND : REAL;
	TIMEBASE : TIME;
	RESET : BOOL;
END_VAR
VAR_OUTPUT
	OUT : REAL;
END_VAR
VAR
	DIFF : REAL;
	OLD_IN : REAL;
	TB : DWORD;
	CET : DWORD;
	CLOCK : TON;
	PROBE : REAL;
END_VAR
END_FUNCTION_BLOCK

(* ---- ROTATION_DIFFERENCE.pou ---- *)
FUNCTION_BLOCK ROTATION_DIFFERENCE
VAR_INPUT
	CURVALUE : UINT;
	LASTVALUE : UINT;
END_VAR
VAR_OUTPUT
	DIFFVALUES : INT;
END_VAR
VAR
	DWCUR : DWORD;
	DWOLD : DWORD;
END_VAR
END_FUNCTION_BLOCK

(* ---- STATISTICS_INT.pou ---- *)
FUNCTION_BLOCK STATISTICS_INT
VAR_INPUT
	IN : INT;
	RESET : BOOL;
END_VAR
VAR_OUTPUT
	MN : INT := 32767;
	MX : INT := -32768;
	AVG : INT;
END_VAR
VAR
	SUM : DINT;
	COUNTER : DINT;
END_VAR
END_FUNCTION_BLOCK

(* ---- STATISTICS_REAL.pou ---- *)
FUNCTION_BLOCK STATISTICS_REAL
VAR_INPUT
	IN : REAL;
	RESET : BOOL;
END_VAR
VAR_OUTPUT
	MN : REAL := 3.402823466E+38;
	MX : REAL := -3.402823466E+38;
	AVG : REAL;
END_VAR
VAR
	COUNTER : DINT;
END_VAR
END_FUNCTION_BLOCK

(* ---- TIMERSWITCH.pou ---- *)
FUNCTION_BLOCK TIMERSWITCH EXTENDS _LConC
VAR_INPUT
	ITFDATETIMEPROVIDER : IDateTimeProvider := Globals.g_dtpDateTimeProvider;
	TCOMPENSATIONSPEED : TIME;
	ASLSCHEDULE : POINTER TO Schedule;
	TZTIMEZONE : REFERENCE TO TimeZone;
END_VAR
VAR_OUTPUT
	EERRORID : ERROR;
	LICLOCKDIFF : LINT;
	EWEEKDAY : WEEKDAY;
	DATTODAY : DATE;
	TODNOW : TIME_OF_DAY;
	STIMEZONE : TZ_NAME;
	EPERIOD : PERIOD;
	DWSWITCHES : DWORD;
END_VAR
VAR
	_LICLOCKSHIFT : LINT;
	_ELASTPERIOD : PERIOD;
	_ULITRANSSTART : ULINT;
	_ULITRANSDURATION : ULINT;
	_PASLSCHEDULE : POINTER TO Schedule;
	_UDIMAXSCHEDULEINDEX : UDINT;
	_PASLHOLIDAYS : POINTER TO Schedule;
	_UDIMAXHOLIDAYSINDEX : UDINT;
	_ULIUTC : ULINT;
	_TZTIMEZONE : TimeZone := TSW.gc_tzTimeZoneCET;
	PTZTIMEZONE : POINTER TO TimeZone;
END_VAR
END_FUNCTION_BLOCK

METHOD CYCLICACTION
VAR_INPUT
	ITFTIMINGCONTROLLER : _ITimingController;
END_VAR
VAR_OUTPUT
	XCOMPLETE : BOOL;
	IERRORID : INT;
END_VAR
END_METHOD

METHOD RESETACTION
VAR_OUTPUT
	XCOMPLETE : BOOL := TRUE;
END_VAR
END_METHOD

METHOD STARTACTION
VAR_OUTPUT
	XCOMPLETE : BOOL := TRUE;
	IERRORID : INT := 0;
END_VAR
END_METHOD

METHOD GETDATETIME : ULINT
VAR_OUTPUT
	EERRORID : ERROR;
END_VAR
END_METHOD

(* ---- UNPACK.pou ---- *)
FUNCTION_BLOCK UNPACK
VAR_INPUT
	B : BYTE;
END_VAR
VAR_OUTPUT
	B0 : BOOL;
	B1 : BOOL;
	B2 : BOOL;
	B3 : BOOL;
	B4 : BOOL;
	B5 : BOOL;
	B6 : BOOL;
	B7 : BOOL;
END_VAR
END_FUNCTION_BLOCK

(* ---- VARIANCE.pou ---- *)
FUNCTION_BLOCK VARIANCE
VAR_INPUT
	IN : REAL;
	RESET : BOOL;
END_VAR
VAR_OUTPUT
	OUT : REAL;
END_VAR
VAR
	Z : DINT;
	A : REAL;
	B : REAL;
END_VAR
END_FUNCTION_BLOCK

(* ---- WORD_AS_BIT.pou ---- *)
FUNCTION_BLOCK WORD_AS_BIT
VAR_INPUT
	W : WORD;
END_VAR
VAR_OUTPUT
	B00 : BOOL;
	B01 : BOOL;
	B02 : BOOL;
	B03 : BOOL;
	B04 : BOOL;
	B05 : BOOL;
	B06 : BOOL;
	B07 : BOOL;
	B08 : BOOL;
	B09 : BOOL;
	B10 : BOOL;
	B11 : BOOL;
	B12 : BOOL;
	B13 : BOOL;
	B14 : BOOL;
	B15 : BOOL;
END_VAR
END_FUNCTION_BLOCK
